// TIA Portal V21 export
// export: Created 2000-01-01T00:00:00.0000000Z, ExportSetting None
VAR_GLOBAL   // PLC tag table "ExchangeTags"
   "电机/运行" AT %M0.0 : Bool;   // 电机运行 / Motor run   {ExternalAccessible false, ExternalWritable false}
   Count AT %MW10 : Word;
END_VAR
VAR_GLOBAL CONSTANT   // user constants
   Limit : Int := 10;
END_VAR
VAR_GLOBAL CONSTANT   // system constants
   LocalModule : Hw_Io := 64;
END_VAR
